// TIA Portal V21 export
Screen "T06_BtnNav"  1024x768, Number=26
  ScreenLayer 
    Button "P_NavBtn" at 0,0 size 100x30  TextOff="BTN", TextOn="BTN"
      EventHandler   EventType=Press
        FunctionCall "ActivateScreen"
          FunctionParameter "Screen name"  Value=Screen_1
